Fanuc KAREL source: kt00503.KL

-- PROVISIONAL review KL for V1013-1; original PC SHA256 f957a0df38d7881cebabed23b3953d5dbe7c553b2739e524bf7a28205105bcf7
-- Incomplete behavior may be omitted. Consult companion uncertainty JSON. Do not deploy.
PROGRAM KT00503
%NOLOCKGROUP
VAR
  OUT : BOOLEAN
-- UNRESOLVED_DECL P1 type=000102
-- UNRESOLVED_DECL P2 type=000106
BEGIN
  -- UNRESOLVED_PC offsets 5-20; opcodes 2E,22,32,35
  -- UNRESOLVED_PC offsets 25-40; opcodes 2E,22,32,35
  -- UNRESOLVED_PC offsets 45-78; opcodes 49,7E,49,7E,AC,23
  -- UNRESOLVED_PC offsets 83-87; opcodes 7F
END KT00503
